SUBAPPLICATION Uebung_094b3f_AX (* Wie Uebung_094b3e_AX, aber ohne T-Stuecke: die Gruppen 1 und 2 sind OptionalGroup_001a bzw. OptionalGroup_002a (Muster mit AOption_IN und AOption_OUT), ihre AOption_OUT speisen AOption_OR_2, dessen OUT die dritte Gruppe OptionalGroup_001b aktiviert. Bei K=1 (DummyGroup) bleibt sie aus. *)
  (* Standard: 61499-2; Description: Copyright (c) 2026 Meisterschulen am Ostbahnhof This program and the accompanying materials are made available under the terms of the Eclipse Public License 2.0 which is available at https://www.eclipse.org/legal/epl-2.0/ SPDX-License-Identifier: EPL-2.0 *)
  (* Version 1.0, 2026-10-17, Franz Höpfinger, Meisterschulen am Ostbahnhof, Kopie von Uebung_094b3_AX, Gruppen 1/2 als OptionalGroup_001a/002a, OR am AOption_OUT, dritte Gruppe 001b. *)
  PACKAGE Uebungen;
  IMPORT Uebungen::const::UT::DefaultPool::InputNumber_I1;
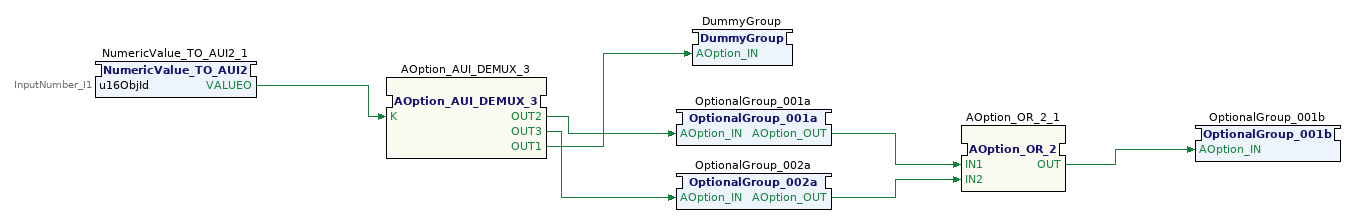
  FBS
    AOption_AUI_DEMUX_3 : Option::selection::AOption_AUI_DEMUX_3;
    AOption_OR_2_1 : Option::merging::AOption_OR_2;
  END_FBS
  SUBAPPS
    NumericValue_TO_AUI2_1 : MyLib::sys::NumericValue_TO_AUI2(u16ObjId := InputNumber_I1);
    OptionalGroup_001a : MyLib_AX_Option::sys::OptionalGroup_001a;
    OptionalGroup_002a : MyLib_AX_Option::sys::OptionalGroup_002a;
    OptionalGroup_001b : MyLib_AX_Option::sys::OptionalGroup_001b;
    DummyGroup : MyLib_AX_Option::sys::DummyGroup;
  END_SUBAPPS
  ADAPTER_CONNECTIONS
    NumericValue_TO_AUI2_1.VALUEO TO AOption_AUI_DEMUX_3.K;
    AOption_AUI_DEMUX_3.OUT2 TO OptionalGroup_001a.AOption_IN;
    AOption_AUI_DEMUX_3.OUT3 TO OptionalGroup_002a.AOption_IN;
    OptionalGroup_001a.AOption_OUT TO AOption_OR_2_1.IN1;
    OptionalGroup_002a.AOption_OUT TO AOption_OR_2_1.IN2;
    AOption_OR_2_1.OUT TO OptionalGroup_001b.AOption_IN;
    AOption_AUI_DEMUX_3.OUT1 TO DummyGroup.AOption_IN;
  END_CONNECTIONS
END_SUBAPPLICATION
